// TIA Portal project "000_empty" (V21)

(* hardware
DEVICE "PLC_1"  S7-1500 station
   slot 0: "Rail_0"  Rack  6ES7 590-1***0-0AA0
   slot 1: "PLC_1"  CPU 1513-1 PN  6ES7 513-1AL02-0AB0  V2.9
      slot 3: "CPU display_1"  6ES7591-1AA00-0AA0
      slot 32768: "PROFINET interface_1"  X1
         slot 32769: "Port_1"  X1 P1
         slot 32770: "Port_2"  X1 P2
      slot 34817: "Virtual CP interface port_1"  Virtual CP interface port  Virtual CP interface port
*)

// ===== PLC "PLC_1"  CPU 1513-1 PN =====

TYPE "UDT_Motor"
   STRUCT
      Running : Bool;   // Motor on
      Speed : Real := 1500.0;   // Speed setpoint
      Count : Int := 7;
   END_STRUCT;
END_TYPE

TYPE "UDT_Inner"
   STRUCT
      Temp : Real := 21.5;
      Input : Bool;
      Static : Int := 3;
      "Return" : DInt;
      Arr : Array[1..3] of Int;
   END_STRUCT;
END_TYPE

TYPE "UDT_Outer"
   STRUCT
      inner : "UDT_Inner";
      innerArr : Array[0..1] of "UDT_Inner";
      s : Struct
         "a" : Bool;
         "m" : Array[0..1, 0..1] of Byte;
      END_STRUCT;
      txt : String[20] := 'outer';
   END_STRUCT;
END_TYPE

DATA_BLOCK "DB_Global"   // DB1
{ S7_Optimized_Access := 'TRUE' }
   VAR
      xBool : Bool := TRUE;   // Bool comment
      iInt : Int := 42;
      rReal : Real := 3.5;   // Real comment
      aInt : Array[0..3] of Int;
      sData : Struct
         "a" : Bool;
         "b" : DInt := -5;
      END_STRUCT;
   END_VAR
BEGIN
   aInt[1] := 11;
END_DATA_BLOCK

DATA_BLOCK "FB_Empty_DB"   // DB2
{ S7_Optimized_Access := 'TRUE' }
VERSION : 0.1
// stored: InstanceOfName FB_Empty
"FB_Empty"
BEGIN
END_DATA_BLOCK

DATA_BLOCK "DB_Motor"   // DB4
{ S7_Optimized_Access := 'TRUE' }
   VAR
      motor : "UDT_Motor";
   END_VAR
BEGIN
   motor.Speed := 750.0;
END_DATA_BLOCK

DATA_BLOCK "FB_Iface_DB"   // DB5
{ S7_Optimized_Access := 'TRUE' }
VERSION : 0.1
// stored: InstanceOfName FB_Iface
"FB_Iface"
BEGIN
   stInt := 99;
   stBool := TRUE;
END_DATA_BLOCK

DATA_BLOCK "DB_AllTypes"   // DB6
{ S7_Optimized_Access := 'TRUE' }
   VAR
      vBool : Bool := TRUE;   // Bool comment
      vByte : Byte := 16#12;
   END_VAR
   VAR RETAIN
      vWord : Word := 16#1234;
   END_VAR
   VAR
      vDWord : DWord := 16#12345678;
      vLWord : LWord := 16#123456789ABCDEF0;
      vSInt : SInt := -12;
      vUSInt : USInt := 200;
      vInt : Int := -1234;
      vUInt : UInt := 60000;
      vDInt : DInt := -123456;
      vUDInt : UDInt := 4000000000;
      vLInt : LInt := -9000000000;
      vULInt : ULInt := 18000000000;
      vReal : Real := 1.5;
      vLReal : LReal := -2.25;
      vS5Time : S5Time := S5T#2S;
      vTime : Time := T#1H2M3S;
      vLTime : LTime := LT#5MS;
      vDate : Date := D#2026-11-05;
      vTod : Time_Of_Day := TOD#12:34:56;
      vLTod : LTime_Of_Day := LTOD#01:02:03.5;
      vDt : Date_And_Time := DT#2026-11-05-12:00:00;
      vLdt : LDT := LDT#2026-11-05-12:00:00;
      vDtl : DTL;
      vChar : Char := 'A';
      vWChar : WChar := WCHAR#'Z';
      vString : String := 'hello';
      vString10 : String[10] := 'ten';
      vWString : WString := WSTRING#'wide';
      vWString5 : WString[5];
      vSetpoint : Int;
      aNeg : Array[-2..2] of Int;
      a2d : Array[0..2, 1..3] of Real;
      a3d : Array[0..1, 0..1, 0..1] of Bool;
      aStr : Array[0..1] of String[8];
      aStruct : Array[0..1] of Struct
         x : Int;
         y : Bool;
      END_STRUCT;
   END_VAR
   VAR RETAIN
      aUdt : Array[0..2] of "UDT_Inner";
   END_VAR
   VAR
      a2dUdt : Array[0..1, 0..1] of "UDT_Outer";
      outer : "UDT_Outer";
      deep : Struct
         l1 : Struct
            l2 : Struct
               v : LReal := 3.14;
               arr : Array[0..1] of Struct
                  z : Word;
               END_STRUCT;
            END_STRUCT;
         END_STRUCT;
      END_STRUCT;
      vTimer : IEC_TIMER;
      vCounter : IEC_COUNTER;
   END_VAR
   VAR RETAIN
      rCount : UDInt;   // Retain counter
      rArr : Array[0..3] of Real;
   END_VAR
BEGIN
   aNeg[-2] := -20;
   aNeg[2] := 20;
   a2d[1,2] := 1.25;
   a3d[1,1,1] := TRUE;
   aStr[1] := 'abc';
   aStruct[1].x := 7;
   a2dUdt[1,0].inner.Static := 5;
   aUdt[2].Temp := 99.5;
   outer.txt := 'changed';
   deep.l1.l2.arr[1].z := 16#BEEF;
   rArr[3] := 0.5;
END_DATA_BLOCK

DATA_BLOCK "DB_NonOpt"   // DB7
{ S7_Optimized_Access := 'FALSE' }
VERSION : 0.1
   VAR
      b0 : Bool;
      b1 : Bool;
      "by" : Byte;
      i : Int := 5;
      d : DInt;
      r : Real;
      t : Time;
      "dt" : Date_And_Time;
      s : String[12] := 'std';
      arr : Array[1..4] of Word;
      "m" : Array[0..1, 0..2] of Int;
      st : Struct
         x : Bool;
         y : Real := 2.5;
      END_STRUCT;
      u : "UDT_Inner";
   END_VAR
BEGIN
   "m"[1,2] := -3;
END_DATA_BLOCK

DATA_BLOCK "DB_OfUdt"   // DB8
{ S7_Optimized_Access := 'TRUE' }
VERSION : 0.1
BEGIN
   txt := 'udtdb';
   inner.Temp := 1.0;
END_DATA_BLOCK

DATA_BLOCK "DB_ArrayDb"   // DB9
{ S7_Optimized_Access := 'TRUE' }
VERSION : 0.1
   VAR
      Header : ArrayDBHeader;
      THIS : Array[0..4] of "UDT_Inner";
   END_VAR
BEGIN
   Header.LowerBound := 0;
   Header.UpperBound := 4;
   Header.Elements := 5;
   Header.PaddedSize := 20;
   Header.ElementSize := 17;
END_DATA_BLOCK

DATA_BLOCK "FB_Multi_DB"   // DB10
{ S7_Optimized_Access := 'TRUE' }
VERSION : 0.1
// stored: InstanceOfName FB_Multi
"FB_Multi"
BEGIN
   cfg.Temp := 30.0;
   mat[1,1] := 11;
   tmrs[2].PT := T#3S;
   sub.stInt := 77;
   subs[1].stInt := 78;
   data.innerArr[1].Arr[2] := 5;
   cnt := 8;
END_DATA_BLOCK

DATA_BLOCK "FB_Top_DB"   // DB11
{ S7_Optimized_Access := 'TRUE' }
VERSION : 0.1
// stored: InstanceOfName FB_Top
"FB_Top"
BEGIN
   "m".sub.stInt := 55;
   ms[0].data.txt := 'deep';
   ms[1].cnt := 9;
END_DATA_BLOCK

DATA_BLOCK "DB_ArrayInt"   // DB12
{ S7_Optimized_Access := 'TRUE' }
VERSION : 0.1
   VAR
      Header : ArrayDBHeader;
      THIS : Array[0..9] of Int;
   END_VAR
BEGIN
   THIS[3] := 33;
   Header.LowerBound := 0;
   Header.UpperBound := 9;
   Header.Elements := 10;
   Header.PaddedSize := 2;
   Header.ElementSize := 2;
END_DATA_BLOCK

// folder: BlockGroup_1

DATA_BLOCK "DB_InGroup"   // DB3
{ S7_Optimized_Access := 'TRUE' }
   VAR
      wWord : Word := 16#00FF;
   END_VAR
BEGIN
END_DATA_BLOCK

// folder: (top level)

FUNCTION_BLOCK "FB_Empty"   // FB1, SCL
{ S7_Optimized_Access := 'TRUE' }
VERSION : 0.1
BEGIN
END_FUNCTION_BLOCK

FUNCTION_BLOCK "FB_Iface"   // FB2, SCL
{ S7_Optimized_Access := 'TRUE' }
VERSION : 0.1
   VAR_INPUT
      iBool : Bool;   // Input bool
      iInt : Int;   // Input int
      iReal : Real;   // Input real
      iArr : Array[0..3] of Int;   // Input array
      iMotor : "UDT_Motor";   // Input UDT
   END_VAR
   VAR_OUTPUT
      oBool : Bool;   // Output bool
      oInt : Int;   // Output int
   END_VAR
   VAR_IN_OUT
      ioReal : Real;   // InOut real
   END_VAR
   VAR
      stInt : Int := 42;   // Static int
      stBool : Bool;   // Static bool comment
   END_VAR
   VAR_TEMP
      tInt : Int;   // Temp int
   END_VAR
   VAR CONSTANT
      cInt : Int := 7;   // Constant int
   END_VAR
BEGIN
   #tInt := #iInt + #cInt;
           #oInt := #tInt;
           #oBool := #iBool;
           #ioReal := #ioReal + #iReal;
END_FUNCTION_BLOCK

FUNCTION_BLOCK "FB_Multi"   // FB3, SCL
{ S7_Optimized_Access := 'TRUE' }
VERSION : 0.1
   VAR_INPUT
      start : Bool;
      cfg : "UDT_Inner";
      mat : Array[0..1, 0..1] of Int;
   END_VAR
   VAR_OUTPUT
      done : Bool;
   END_VAR
   VAR_IN_OUT
      io : Real;
   END_VAR
   VAR
      tmr : TON_TIME;
      tmrs : Array[0..2] of TON_TIME;
      ctr : CTU_INT;
      edge : R_TRIG;
      sub : "FB_Iface";
      subs : Array[0..1] of "FB_Iface";
      data : "UDT_Outer";
      cnt : Int := 4;
      Temp : Int;
   END_VAR
   VAR RETAIN
      r1 : Int := 6;
      r2 : Real;
   END_VAR
   VAR_TEMP
      t1 : Int;
   END_VAR
BEGIN
   #tmr(IN := #start, PT := T#1S);
           #done := #tmr.Q;
END_FUNCTION_BLOCK

FUNCTION_BLOCK "FB_Top"   // FB4, SCL
{ S7_Optimized_Access := 'TRUE' }
VERSION : 0.1
   VAR
      "m" : "FB_Multi";
      ms : Array[0..1] of "FB_Multi";
      x : Real;
   END_VAR
BEGIN
   #m(start := TRUE, io := #x);
END_FUNCTION_BLOCK

ORGANIZATION_BLOCK "Main"   // OB1, LAD, ProgramCycle
TITLE = "Main Program Sweep (Cycle)"
{ S7_Optimized_Access := 'TRUE' }
VERSION : 0.1
   VAR_INPUT
      Initial_Call : Bool;   // Initial call of this OB
      Remanence : Bool;   // =True, if remanent data are available
   END_VAR
BEGIN
END_ORGANIZATION_BLOCK